DATA_BLOCK "FRK_PersistStatus"
{ S7_Optimized_Access := 'TRUE' }
VERSION : 0.1
NON_RETAIN
VAR
    SchemaVersion {ExternalWritable := 'False'} : UInt := 1;
    Medium {ExternalWritable := 'False'} : String[16] := 'LOAD_DB';
    Restoring {ExternalWritable := 'False'} : Bool;
    Failed {ExternalWritable := 'False'} : Bool;
    NativeStatus {ExternalWritable := 'False'} : Word;
    DocumentCount {ExternalWritable := 'False'} : Int := 20;
END_VAR
BEGIN
END_DATA_BLOCK
